FUNCTION_BLOCK CMoGetLocalDateTime
VAR_INPUT
END_VAR
VAR_OUTPUT
END_VAR
VAR_IN_OUT
    DateTime        : CMoDateTime;
END_VAR
VAR
	fbLocalTime     : FB_LocalSystemTime := (bEnable := TRUE, dwCycle := 1);
END_VAR

// =============================================================================
// CMoGetLocalDateTime — Read Local System Time (Beckhoff)
// CMo Library v1.0
// Requires: Tc2_Utilities library
// =============================================================================
// Reads the local Windows system time via FB_LocalSystemTime and
// maps TIMESTRUCT fields into CMoDateTime.
//
// Must be called cyclically. Called internally by CMoMainRuntime
// every scan.
//
// Usage:
//   fbLocal(DateTime := Framework.CurrentLocalDateTime);
// =============================================================================

fbLocalTime();
IF fbLocalTime.bValid THEN
    DateTime.Year        := WORD_TO_DINT(fbLocalTime.systemTime.wYear);
    DateTime.Month       := WORD_TO_DINT(fbLocalTime.systemTime.wMonth);
    DateTime.Day         := WORD_TO_DINT(fbLocalTime.systemTime.wDay);
    DateTime.Hour        := WORD_TO_DINT(fbLocalTime.systemTime.wHour);
    DateTime.Minute      := WORD_TO_DINT(fbLocalTime.systemTime.wMinute);
    DateTime.Second      := WORD_TO_DINT(fbLocalTime.systemTime.wSecond);
    DateTime.MicroSecond := WORD_TO_DINT(fbLocalTime.systemTime.wMilliseconds) * 1000;
    DateTime.IsLocal     := TRUE;
END_IF;

END_FUNCTION_BLOCK

(* stored: Version 1.1.0.1, ProductVersion 3.1.4024.16
   POU CMoGetLocalDateTime: Id {8cb8b7b6-173d-45a1-9618-7b1cf0721494}, SpecialFunc None *)
